SUBAPPLICATION Uebung_266_AX (* Dimmer am Terminal: wie 265, zusaetzlich Softkey F1 als zweite Bedienstelle (tippen = ein/aus, halten = dimmen) und Helligkeit in % auf OutputNumber_N1 *)
  (* Standard: 61499-2; Description: Copyright (c) 2026 Meisterschulen am Ostbahnhof This program and the accompanying materials are made available under the terms of the Eclipse Public License 2.0 which is available at https://www.eclipse.org/legal/epl-2.0/ SPDX-License-Identifier: EPL-2.0 *)
  (* Version 1.0, 2026-11-07, Franz Höpfinger, Meisterschulen am Ostbahnhof, initial API and implementation and/or initial documentation *)
  PACKAGE Uebungen;
  IMPORT logiBUS::io::DI::logiBUS_DI::Input_I1;
  IMPORT logiBUS::io::DI::logiBUS_DI::Input_I2;
  IMPORT logiBUS::io::DI::logiBUS_DI::Input_I3;
  IMPORT logiBUS::io::DI::logiBUS_DI_Events::BUTTON_LONG_PRESS_START;
  IMPORT logiBUS::io::DI::logiBUS_DI_Events::BUTTON_LONG_PRESS_UP;
  IMPORT logiBUS::io::DI::logiBUS_DI_Events::BUTTON_SINGLE_CLICK;
  IMPORT logiBUS::io::DQ::logiBUS_DO::Output_Q1;
  IMPORT Uebungen::const::UT::DefaultPool::OutputNumber_N1;
  IMPORT Uebungen::const::UT::DefaultPool::SoftKey_F1;
  IMPORT isobus::UT::io::Softkey::SoftKeyActivationCode::SK_RELEASED;
  IMPORT isobus::UT::io::Softkey::SoftKeyActivationCode::SK_STILL_HELD_START;
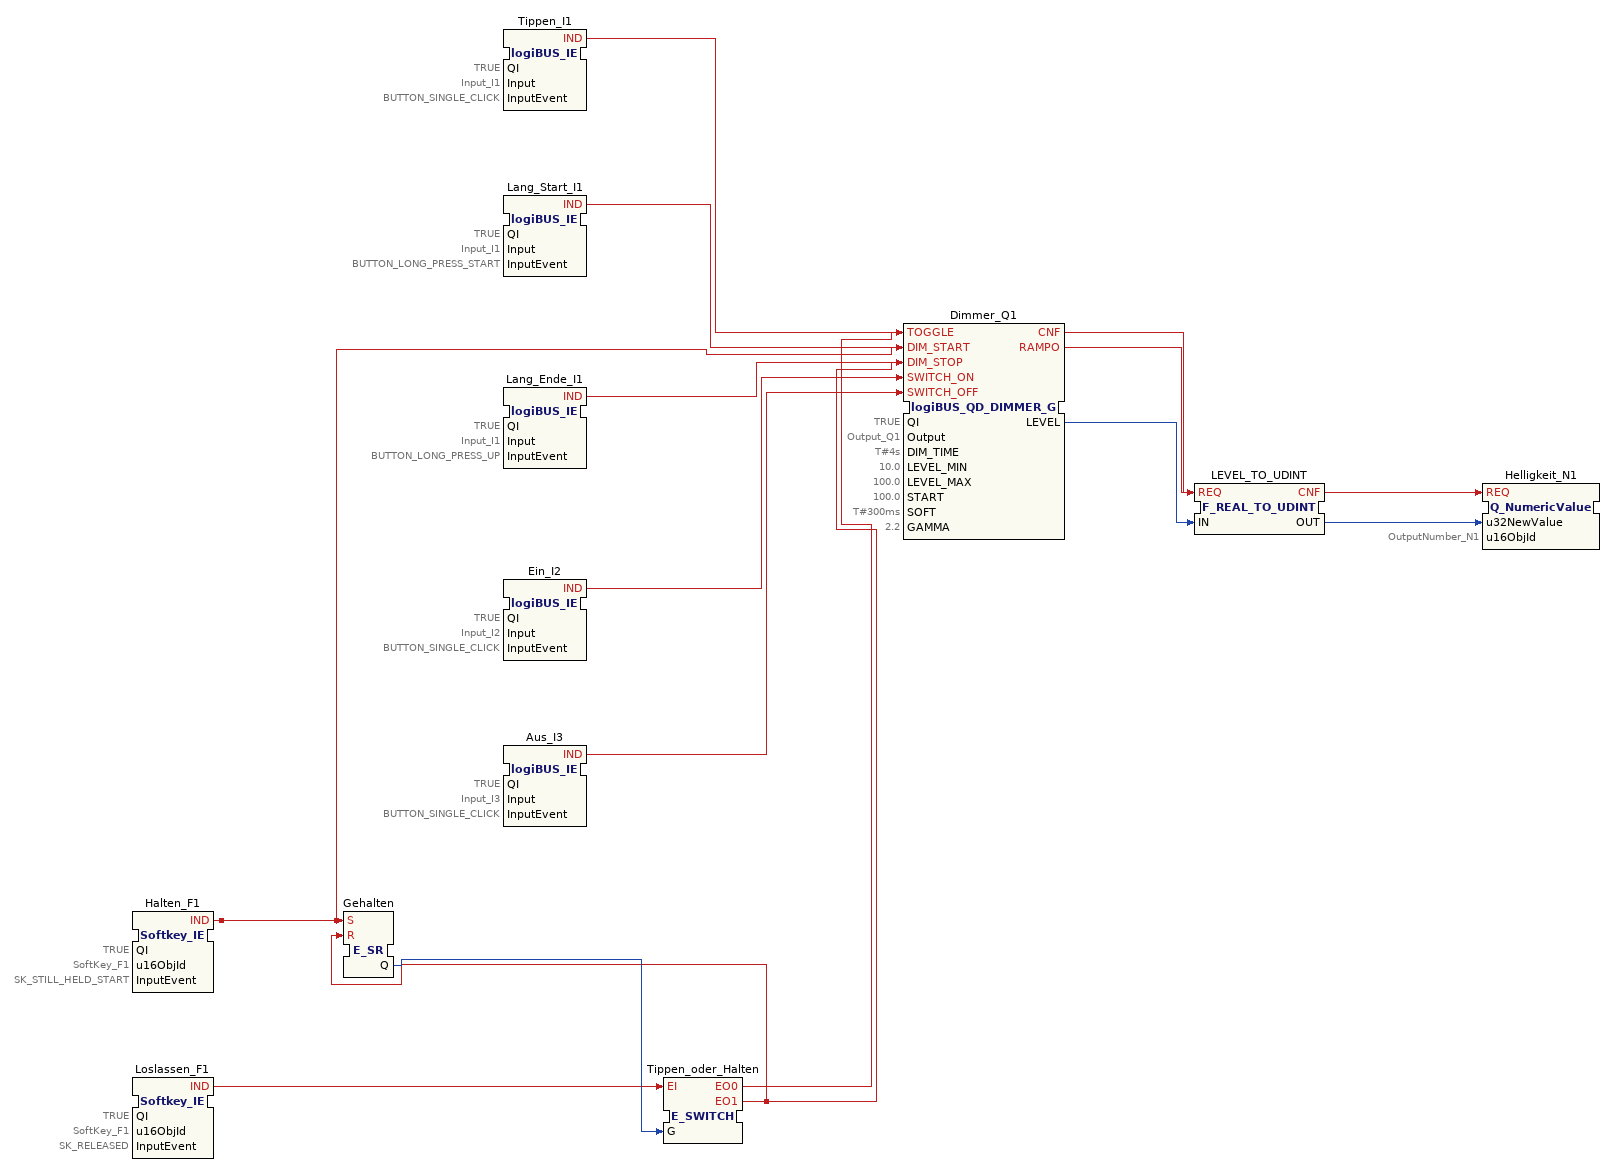
  FBS
    Tippen_I1 : logiBUS::io::DI::logiBUS_IE(QI := TRUE, Input := Input_I1, InputEvent := BUTTON_SINGLE_CLICK);
    Lang_Start_I1 : logiBUS::io::DI::logiBUS_IE(QI := TRUE, Input := Input_I1, InputEvent := BUTTON_LONG_PRESS_START);
    Lang_Ende_I1 : logiBUS::io::DI::logiBUS_IE(QI := TRUE, Input := Input_I1, InputEvent := BUTTON_LONG_PRESS_UP);
    Ein_I2 : logiBUS::io::DI::logiBUS_IE(QI := TRUE, Input := Input_I2, InputEvent := BUTTON_SINGLE_CLICK);
    Aus_I3 : logiBUS::io::DI::logiBUS_IE(QI := TRUE, Input := Input_I3, InputEvent := BUTTON_SINGLE_CLICK);
    Halten_F1 : isobus::UT::io::Softkey::Softkey_IE(QI := TRUE, u16ObjId := SoftKey_F1, InputEvent := SK_STILL_HELD_START);
    Loslassen_F1 : isobus::UT::io::Softkey::Softkey_IE(QI := TRUE, u16ObjId := SoftKey_F1, InputEvent := SK_RELEASED);
    Gehalten : iec61499::events::E_SR;
    Tippen_oder_Halten : iec61499::events::E_SWITCH;
    Dimmer_Q1 : logiBUS::io::DQ::logiBUS_QD_DIMMER_G(QI := TRUE, Output := Output_Q1, DIM_TIME := T#4s, LEVEL_MIN := 10.0, LEVEL_MAX := 100.0, START := 100.0, SOFT := T#300ms, GAMMA := 2.2);
    LEVEL_TO_UDINT : iec61131::conversion::F_REAL_TO_UDINT;
    Helligkeit_N1 : isobus::UT::Q::Q_NumericValue(u16ObjId := OutputNumber_N1);
  END_FBS
  EVENT_CONNECTIONS
    Tippen_I1.IND TO Dimmer_Q1.TOGGLE;
    Lang_Start_I1.IND TO Dimmer_Q1.DIM_START;
    Lang_Ende_I1.IND TO Dimmer_Q1.DIM_STOP;
    Ein_I2.IND TO Dimmer_Q1.SWITCH_ON;
    Aus_I3.IND TO Dimmer_Q1.SWITCH_OFF;
    Halten_F1.IND TO Gehalten.S;
    Halten_F1.IND TO Dimmer_Q1.DIM_START;
    Loslassen_F1.IND TO Tippen_oder_Halten.EI;
    Tippen_oder_Halten.EO0 TO Dimmer_Q1.TOGGLE;
    Tippen_oder_Halten.EO1 TO Dimmer_Q1.DIM_STOP;
    Tippen_oder_Halten.EO1 TO Gehalten.R;
    Dimmer_Q1.CNF TO LEVEL_TO_UDINT.REQ;
    Dimmer_Q1.RAMPO TO LEVEL_TO_UDINT.REQ;
    LEVEL_TO_UDINT.CNF TO Helligkeit_N1.REQ;
  END_CONNECTIONS
  DATA_CONNECTIONS
    Gehalten.Q TO Tippen_oder_Halten.G;
    Dimmer_Q1.LEVEL TO LEVEL_TO_UDINT.IN;
    LEVEL_TO_UDINT.OUT TO Helligkeit_N1.u32NewValue;
  END_CONNECTIONS
END_SUBAPPLICATION
